(* IEC 61131-3 sources: iecf/harness/cases/codesysmembershadow.d, 1 file *)

(* ---- lib.st ---- *)
FUNCTION_BLOCK StopTask
  VAR_OUTPUT q : INT; END_VAR
  q := 1000;
END_FUNCTION_BLOCK

FUNCTION Helper : INT
  Helper := 1000;
END_FUNCTION

FUNCTION Twice : INT
  VAR_INPUT x : INT; END_VAR
  Twice := 2 * x;
END_FUNCTION
